(* PLC project g_phase_hold_permissive_bomb, Anonymous Benchmark Suite 1.0 *)
(* stored: creationDateTime 2026-09-02T00:00:00 *)

PROGRAM g_phase_hold_permissive_bomb
  VAR_INPUT
    run_command : BOOL;
    agitator_ok : BOOL;
    resume_command : BOOL;
    maint : BOOL;
  END_VAR
  VAR_OUTPUT
    held : BOOL;
    heater : BOOL;
  END_VAR

(* LD diagram, written out as Structured Text *)
held := run_command AND NOT agitator_ok OR held AND NOT resume_command;
heater := run_command AND NOT held AND agitator_ok OR held AND maint;
END_PROGRAM

CONFIGURATION Config0
  RESOURCE Res0 ON PLC
    TASK tcyclic(INTERVAL := T#10ms, PRIORITY := 0);
    PROGRAM inst0 WITH tcyclic : g_phase_hold_permissive_bomb;
  END_RESOURCE
END_CONFIGURATION
